(* IEC 61131-3 sources: SRCI_CLIENT_PLC/RobotLibrary/Library/POUs/Spline/MC_CreateSpline/Structures, 4 files *)

(* ---- CreateSplineOutCmd.st ---- *)
{attribute 'pack_mode' := '1'}
// -------------------------------------------------------------------------
//  SRCI Robot Library
// -------------------------------------------------------------------------
//
//  Object:      CreateSplineOutCmd
//  Author:      Thorsten Brach
//  Date:        2024-08-01
//
//  Description:
//
//
//  Copyright:
//    (C) 2024 Thorsten Brach. All rights reserved
//             Licensed under the MIT License.
//
//  Disclaimer:
//    This project is provided without any guarantee and can be used for
//    private and commercial purposes. Any use is at the user’s
//    own risk and responsibility.
//
// -------------------------------------------------------------------------
TYPE CreateSplineOutCmd :
STRUCT
END_STRUCT
END_TYPE

(* ---- CreateSplineParCmd.st ---- *)
{attribute 'pack_mode' := '1'}
// -------------------------------------------------------------------------
//  SRCI Robot Library
// -------------------------------------------------------------------------
//
//  Object:      CreateSplineParCmd
//  Author:      Thorsten Brach
//  Date:        2024-08-01
//
//  Description:
//
//
//  Copyright:
//    (C) 2024 Thorsten Brach. All rights reserved
//             Licensed under the MIT License.
//
//  Disclaimer:
//    This project is provided without any guarantee and can be used for
//    private and commercial purposes. Any use is at the user’s
//    own risk and responsibility.
//
// -------------------------------------------------------------------------
TYPE CreateSplineParCmd :
STRUCT
  /// Define the method to calculate the path trajectory for the spline movement
  Mode            : SplineMode;
  /// Index of the spline trajectory to be created
  SplineID        : SINT;
  /// Contains all data relevant to the spline trajectory
  /// • Cartesian position
  /// • Coordinate systems
  /// • Dynamic parameters
  /// For more information refer to chapter 5.5.13.3
  SplineData      : ARRAY[1..RobotLibraryParameter.SPLINE_DATA_MAX] OF SplineData;
END_STRUCT
END_TYPE

(* ---- CreateSplineRecvData.st ---- *)
{attribute 'pack_mode' := '1'}
// -------------------------------------------------------------------------
//  SRCI Robot Library
// -------------------------------------------------------------------------
//
//  Object:      CreateSplineRecvData
//  Author:      Thorsten Brach
//  Date:        2024-08-01
//
//  Description:
//
//
//  Copyright:
//    (C) 2024 Thorsten Brach. All rights reserved
//             Licensed under the MIT License.
//
//  Disclaimer:
//    This project is provided without any guarantee and can be used for
//    private and commercial purposes. Any use is at the user’s
//    own risk and responsibility.
//
// -------------------------------------------------------------------------
TYPE CreateSplineRecvData EXTENDS RspHeader :
STRUCT
END_STRUCT
END_TYPE

(* ---- CreateSplineSendData.st ---- *)
{attribute 'pack_mode' := '1'}
// -------------------------------------------------------------------------
//  SRCI Robot Library
// -------------------------------------------------------------------------
//
//  Object:      CreateSplineSendData
//  Author:      Thorsten Brach
//  Date:        2024-08-01
//
//  Description:
//
//
//  Copyright:
//    (C) 2024 Thorsten Brach. All rights reserved
//             Licensed under the MIT License.
//
//  Disclaimer:
//    This project is provided without any guarantee and can be used for
//    private and commercial purposes. Any use is at the user’s
//    own risk and responsibility.
//
// -------------------------------------------------------------------------
TYPE CreateSplineSendData EXTENDS CmdHeader:
STRUCT
  /// Define the method to calculate the path trajectory for the spline movement
  Mode            : UINT;
  /// Index of the spline trajectory to be created
  SplineID        : SINT;
  /// Contains all data relevant to the spline trajectory
  /// • Cartesian position
  /// • Coordinate systems
  /// • Dynamic parameters
  /// For more information refer to chapter 5.5.13.3
  SplineData      : ARRAY[1..RobotLibraryParameter.SPLINE_DATA_MAX] OF SplineDataSend;
END_STRUCT
END_TYPE
